ABB RobotStudio station: Pallet_Project.rspag

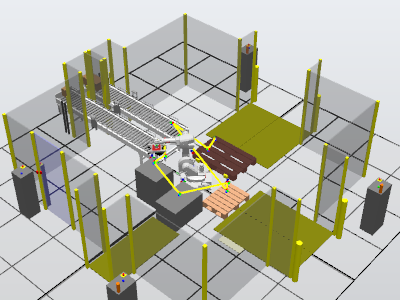
--- station ---
Station Pallet_Project (saved by RobotStudio 25.2.11220.0)
Controller Controler
  mechanical unit ROB_1: IRB1600_10_145__02, 6 joints, base frame (0, 0, 0) mm, rotated rx 0 ry 0 rz 135 deg
Layout (positions relative to the parent item):
  - IRB1600_10_145__02 [mechanism, from %ABB.RobotStudio.Models.IRB1600%\IRB1600_10_145_G_02.rslib] at (0, 0, 0) mm, rotated rx 0 ry 0 rz 135 deg; joint values [0, 0, 0, 0, 1.5708, 0] (rad or m)
  - Half EPAL [part] at (-400, -600, 0) mm, rotated rx 0 ry 0 rz -90 deg, size 600 x 800 x 144 mm
  - ConveyorBox1 [part, from %ABB.RobotStudio.Models.Conveyors%\Conveyor Guide 400.rslib] at (150, 3660, 0) mm, rotated rx 0 ry 0 rz -90 deg
  - ConveyorBox2 [part, from %ABB.RobotStudio.Models.Conveyors%\Conveyor Guide 400.rslib] at (-550, 3660, 0) mm, rotated rx 0 ry 0 rz -90 deg
  - PalletizingVacuumTool [mechanism] at (-530.33, 530.33, 1121.5) mm, rotated rx 180 ry 0 rz -45 deg
      TCP toolVacuum at (0, 0, 175) mm
      links: PalletizingVacuumTool
  - Box1 [part] at (338.5, 3410, 868) mm, size 249 x 499 x 200 mm
  - Box2 [part] at (-353.5, 3575, 868) mm, size 129 x 129 x 200 mm
  - EuroPallet [part, from Components\EuroPalletWood.rslib] at (1400, -600, 0) mm, rotated rx 0 ry 0 rz 90 deg
  - StackingTable [part], size 500 x 600 x 770 mm
  - LinerStand [part], size 800 x 540 x 500 mm
  - SC_Conveyor1 [smart component]
      signals: DO BoxArrived, DI EuroPalletReplaced, DO EuroPalletReplacedOut, DI EuroPalletFull
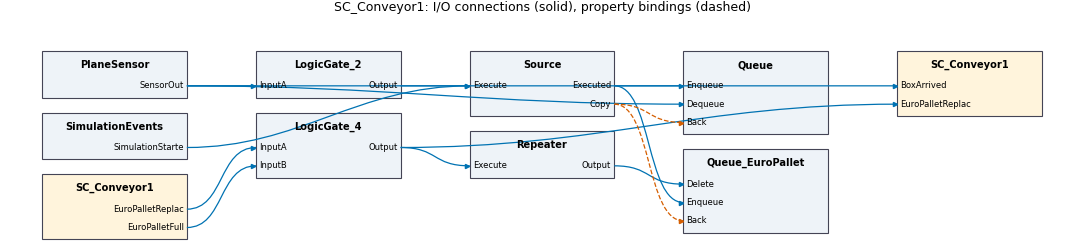
      connections:
        Source.Executed -> Queue.Enqueue
        PlaneSensor.SensorOut -> Queue.Dequeue
        PlaneSensor.SensorOut -> SC_Conveyor1.BoxArrived
        PlaneSensor.SensorOut -> LogicGate_2.InputA
        LogicGate_2.Output -> Source.Execute
        SimulationEvents.SimulationStarted -> Source.Execute
        SC_Conveyor1.EuroPalletReplaced -> LogicGate_4.InputA
        SC_Conveyor1.EuroPalletFull -> LogicGate_4.InputB
        LogicGate_4.Output -> SC_Conveyor1.EuroPalletReplacedOut
        LogicGate_4.Output -> Repeater.Execute
        Repeater.Output -> Queue_EuroPallet.Delete
        Source.Executed -> Queue_EuroPallet.Enqueue
        Source.Copy => Queue.Back
        Source.Copy => Queue_EuroPallet.Back
    - Source [smart component, from Components\Source.rslib]
        properties: Source=Box1; Copy=(none); Parent=(none); Position=[0.3385 3.39 0.868]; Orientation=[0 0 0]; Transient=true; PhysicsBehavior=-1
    - Queue [smart component, from Components\Queue.rslib]
        properties: Back=(none); Front=(none); Queue={70ca05b0-7144-4f49-83d8-d915b94a0a02};{7705e30e-55ab-4cc9-9220-690ff83121bf};{02bf6a2a-9363-4f0e-8f48-ba3ac55a3133};{2a754624-700a-40ce-a7f5-ac92a5654210};{9528570a-eb81-4ef3-89d0-eb89feb3dc99};{56097831-269e-4b26-b9dc-fc2a065cc4d2};{84102578-6d50-4318-bba9-f08da63948c5};{ab344251-b794-483f-853d-2cd57e9333d1};{43a68e49-bc40-4bf4-a0b0-52db603239fa};{90f7df2a-bd47-43a1-93ae-0975fdea56be};{8df4c4d2-3a0e-4db8-a3f9-2112c5fdeae1};{a6db4b97-f991-4390-b4fd-8137cccb983c};{ac275fb4-aa41-4d4d-8111-4fbb0763e808}; NumberOfObjects=1
    - LinearMover [smart component, from Components\LinearMover.rslib]
        properties: Object=Queue; Direction=[0 -0.001 0]; Speed=0.25; Reference=Global; ReferenceObject=(none)
    - PlaneSensor [smart component, from Components\PlaneSensor.rslib]
        properties: Origin=[0.1885 0.675 0.788]; Axis1=[0.3 0 0]; Axis2=[0 0 0.01]; Tag=(none); SenseMultiple=false; SensedPart=(none)
      - _sensorPart_ [part], size 300 x 0 x 10 mm
    - LogicGate_2 [smart component, from Components\LogicGate.rslib]
        properties: Operator=NOT; Delay=0
    - SimulationEvents [smart component, from Components\SimulationEvents.rslib]
    - Queue_EuroPallet [smart component, from Components\Queue.rslib]
        properties: Back=(none); Front=(none); Queue=; NumberOfObjects=0
    - LogicGate_4 [smart component, from Components\LogicGate.rslib]
        properties: Operator=AND; Delay=0
    - Repeater [smart component, from Components\Repeater.rslib]
        properties: Count=12
  - SC_Gripper [smart component]
      signals: DI Grip
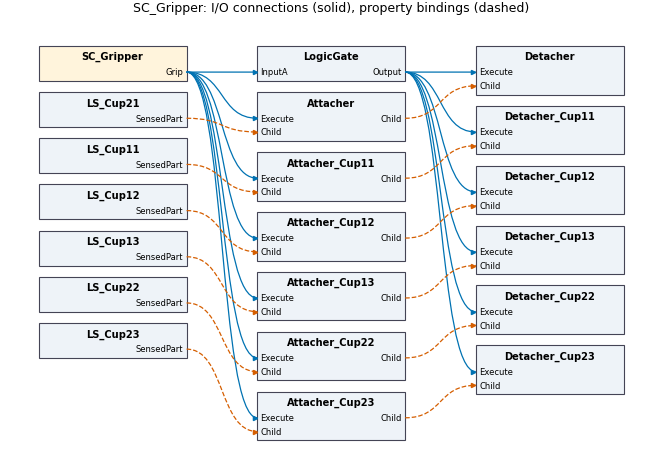
      connections:
        SC_Gripper.Grip -> Attacher.Execute
        SC_Gripper.Grip -> LogicGate.InputA
        LogicGate.Output -> Detacher.Execute
        SC_Gripper.Grip -> Attacher_Cup11.Execute
        LogicGate.Output -> Detacher_Cup11.Execute
        SC_Gripper.Grip -> Attacher_Cup12.Execute
        LogicGate.Output -> Detacher_Cup12.Execute
        SC_Gripper.Grip -> Attacher_Cup13.Execute
        LogicGate.Output -> Detacher_Cup13.Execute
        SC_Gripper.Grip -> Attacher_Cup22.Execute
        LogicGate.Output -> Detacher_Cup22.Execute
        SC_Gripper.Grip -> Attacher_Cup23.Execute
        LogicGate.Output -> Detacher_Cup23.Execute
        LS_Cup21.SensedPart => Attacher.Child
        Attacher.Child => Detacher.Child
        LS_Cup11.SensedPart => Attacher_Cup11.Child
        Attacher_Cup11.Child => Detacher_Cup11.Child
        LS_Cup12.SensedPart => Attacher_Cup12.Child
        Attacher_Cup12.Child => Detacher_Cup12.Child
        LS_Cup13.SensedPart => Attacher_Cup13.Child
        Attacher_Cup13.Child => Detacher_Cup13.Child
        LS_Cup22.SensedPart => Attacher_Cup22.Child
        Attacher_Cup22.Child => Detacher_Cup22.Child
        LS_Cup23.SensedPart => Attacher_Cup23.Child
        Attacher_Cup23.Child => Detacher_Cup23.Child
    - LS_Cup21 [smart component, from Components\LineSensor.rslib] at (0, 0, 0) mm
        properties: Start=[-0.597509982704304 0.689429996191639 0.956499992313755]; End=[-0.597509981617333 0.689429995104668 0.924499992313755]; Length=0.032; Radius=0.00331491712707182; Tag=(none); SenseMultiple=false; SensedPart=(none); SensedPoint=[0 0 0]
      - _sensorPart_ [part], size 6.4 x 6.4 x 32 mm
    - Attacher [smart component, from Components\Attacher.rslib]
        properties: Parent=PalletizingVacuumTool; Flange=0; Child=(none); Mount=false; Offset=[0 0 0]; Orientation=[0 0 0]
    - Detacher [smart component, from Components\Detacher.rslib]
        properties: Child=(none); KeepPosition=true
    - LogicGate [smart component, from Components\LogicGate.rslib]
        properties: Operator=NOT; Delay=0
    - LS_Cup11 [smart component, from Components\LineSensor.rslib]
        properties: Start=[-0.68943 0.59751 0.9565]; End=[-0.68943 0.59751 0.9245]; Length=0.032; Radius=0.00331; Tag=(none); SenseMultiple=false; SensedPart=(none); SensedPoint=[0 0 0]
      - _sensorPart_ [part], size 6.6 x 6.6 x 32 mm
    - LS_Cup12 [smart component, from Components\LineSensor.rslib]
        properties: Start=[-0.57629 0.48437 0.9565]; End=[-0.57629 0.48437 0.9245]; Length=0.032; Radius=0.00331; Tag=(none); SenseMultiple=false; SensedPart=(none); SensedPoint=[0 0 0]
      - _sensorPart_ [part], size 6.6 x 6.6 x 32 mm
    - LS_Cup13 [smart component, from Components\LineSensor.rslib]
        properties: Start=[-0.46315 0.37123 0.9565]; End=[-0.46315 0.37123 0.9245]; Length=0.032; Radius=0.00331; Tag=(none); SenseMultiple=false; SensedPart=(none); SensedPoint=[0 0 0]
      - _sensorPart_ [part], size 6.6 x 6.6 x 32 mm
    - LS_Cup22 [smart component, from Components\LineSensor.rslib]
        properties: Start=[-0.48437 0.57629 0.9565]; End=[-0.48437 0.57629 0.9245]; Length=0.032; Radius=0.00331; Tag=(none); SenseMultiple=false; SensedPart=(none); SensedPoint=[0 0 0]
      - _sensorPart_ [part], size 6.6 x 6.6 x 32 mm
    - LS_Cup23 [smart component, from Components\LineSensor.rslib]
        properties: Start=[-0.37123 0.46315 0.9565]; End=[-0.37123 0.46315 0.9245]; Length=0.032; Radius=0.00331; Tag=(none); SenseMultiple=false; SensedPart=(none); SensedPoint=[0 0 0]
      - _sensorPart_ [part], size 6.6 x 6.6 x 32 mm
    - Attacher_Cup11 [smart component, from Components\Attacher.rslib]
        properties: Parent=PalletizingVacuumTool; Flange=0; Child=(none); Mount=false; Offset=[0 0 0]; Orientation=[0 0 0]
    - Detacher_Cup11 [smart component, from Components\Detacher.rslib]
        properties: Child=(none); KeepPosition=true
    - Attacher_Cup12 [smart component, from Components\Attacher.rslib]
        properties: Parent=PalletizingVacuumTool; Flange=0; Child=(none); Mount=false; Offset=[0 0 0]; Orientation=[0 0 0]
    - Detacher_Cup12 [smart component, from Components\Detacher.rslib]
        properties: Child=(none); KeepPosition=true
    - Attacher_Cup13 [smart component, from Components\Attacher.rslib]
        properties: Parent=PalletizingVacuumTool; Flange=0; Child=(none); Mount=false; Offset=[0 0 0]; Orientation=[0 0 0]
    - Detacher_Cup13 [smart component, from Components\Detacher.rslib]
        properties: Child=(none); KeepPosition=true
    - Attacher_Cup22 [smart component, from Components\Attacher.rslib]
        properties: Parent=PalletizingVacuumTool; Flange=0; Child=(none); Mount=false; Offset=[0 0 0]; Orientation=[0 0 0]
    - Detacher_Cup22 [smart component, from Components\Detacher.rslib]
        properties: Child=(none); KeepPosition=true
    - Attacher_Cup23 [smart component, from Components\Attacher.rslib]
        properties: Parent=PalletizingVacuumTool; Flange=0; Child=(none); Mount=false; Offset=[0 0 0]; Orientation=[0 0 0]
    - Detacher_Cup23 [smart component, from Components\Detacher.rslib]
        properties: Child=(none); KeepPosition=true
  - SC_Conveyor2 [smart component]
      signals: DO BoxArrived, DI HalfPalletReplaced, DI HalfPalletFull, DO HalfPalletReplacedOut
      connections:
        Source.Executed -> Queue.Enqueue
        PlaneSensor.SensorOut -> Queue.Dequeue
        PlaneSensor.SensorOut -> SC_Conveyor2.BoxArrived
        PlaneSensor.SensorOut -> LogicGate.InputA
        SimulationEvents.SimulationStarted -> Source.Execute
        Source.Executed -> Queue_HalfPallet.Enqueue
        LogicGate.Output -> Source.Execute
        Repeater.Output -> Queue_HalfPallet.Delete
        SC_Conveyor2.HalfPalletReplaced -> LogicGate_5.InputA
        SC_Conveyor2.HalfPalletFull -> LogicGate_5.InputB
        LogicGate_5.Output -> Repeater.Execute
        LogicGate_5.Output -> SC_Conveyor2.HalfPalletReplacedOut
        Source.Copy => Queue.Back
        Source.Copy => Queue_HalfPallet.Back
    - Source [smart component, from Components\Source.rslib]
        properties: Source=Box2; Copy=(none); Parent=(none); Position=[-0.3535 3.575 0.868]; Orientation=[0 0 0]; Transient=true; PhysicsBehavior=-1
    - Queue [smart component, from Components\Queue.rslib]
        properties: Back=(none); Front=(none); Queue={648eb2a2-8d13-4a50-a9a9-4bb0657455f7};{41be35e7-4a03-4cb4-92d6-970da98b32eb};{4f5e8617-4ef4-4248-bc63-4e8ec75bf0fd};{9850fa1d-30e0-46cb-a9aa-89d687d5a572};{8673d542-8e4c-49b3-88b3-ba839af60b27};{121a61d2-9307-4f78-a061-101ab78a5607};{316e579a-2297-4da1-921e-c195e3c1eac9};{afd6ccd5-80c3-46f0-a33f-b3bd5f1b0761};{a691a1e4-6464-4329-bb8e-435514d80af1};{358ac2eb-a4d6-456f-aa39-476db23d4f48}; NumberOfObjects=1
    - LinearMover [smart component, from Components\LinearMover.rslib]
        properties: Object=Queue; Direction=[0 -0.001 0]; Speed=0.25; Reference=Global; ReferenceObject=(none)
    - PlaneSensor [smart component, from Components\PlaneSensor.rslib]
        properties: Origin=[-0.5035 0.675 0.788]; Axis1=[0.3 0 0]; Axis2=[0 0 0.01]; Tag=(none); SenseMultiple=false; SensedPart=(none)
      - _sensorPart_ [part], size 300 x 0 x 10 mm
    - LogicGate [smart component, from Components\LogicGate.rslib]
        properties: Operator=NOT; Delay=0
    - SimulationEvents [smart component, from Components\SimulationEvents.rslib]
    - Queue_HalfPallet [smart component, from Components\Queue.rslib]
        properties: Back=(none); Front=(none); Queue={f5edb1ce-3bf5-426a-a389-0b0047efa949};{5ce0816a-b692-43c6-82f7-492eb3fc1c7c};{ad3ef4b5-2c59-4daa-9658-0c77e5efb67d};{c9c476d0-74ff-4b18-bfb3-2d6c852b8493};{1bf865c6-1649-4319-b5ff-cd81faaa6069};{f626778c-15a6-4059-b27a-7c8f9da4f34f};{a60dd0dd-490e-48fe-bb32-16f415136b44};{4ec9b3b2-e4a8-4d14-aea0-9552a35d2afd};{38bc6a68-8d9e-44a7-a5f0-badb214ea710};{f9543542-377a-43f1-9613-018dced76680};{486b4c2f-b225-4486-b430-5ab7d813c599};{7da52d9e-9053-4b1a-839c-0aedc5495cc7};{c2400356-fde5-4523-9dc7-d26788098951};{75099568-1fe6-4c34-8328-63fd42144c3b};{8ca6c374-2d39-4938-8324-38c48ae4f51d};{f3c160ab-6f5f-460b-8b54-c2c3b0bc175f};{1c289510-9a29-4e1c-b603-54b7a0027260};{d39da69b-e59a-4ace-85a5-bba54583b01c};{bc328c62-4bf3-4a57-965c-0c93e0ee296d};{60f4dcb3-d366-4d0b-b05a-5b2073fcd9e8};{44334a49-cf52-4d95-9964-3bb568ce732d};{f9240695-1965-47e5-bcd4-644ec5904899};{72a970fd-f238-4ac5-b811-00686975bc20};{bd297b2a-4ad7-44fa-87c8-1ac40b0d2fbf};{3dafa88d-62b0-429f-9c75-c8c7bde09fc6};{a7d8f176-4e9d-4819-8805-982bee0c310d};{72ae6bb6-3373-4f60-a321-dfdc0981c562};{fff16105-3d56-4b21-a888-399904fd95d4};{56e4abf9-acd4-4a00-b067-52a58200d221};{2eb8ae55-b553-4f83-b65d-07c27c701dd6};{dfb05241-1220-45e8-b584-1559777c0125};{49a2c23a-27ea-4b0b-af5c-f9d01014f642};{0adfb5d7-4fd0-41be-8361-c42c9d28ca51};{8cf74624-f46b-49ca-a524-038ddb88ba0f};{bde2cdc4-b3e4-48fe-8333-d64185b5a8e7};{d17564c2-89d4-4b4f-8596-5dca9165a286};{6fec26e7-cb1b-4d74-b4a6-8ed7a2eb81a6};{e04d8697-cc19-4df5-b7fa-dff41516820c};{134714af-70a5-49a3-8b99-ea847d1ef329};{23aa8eff-aaeb-4079-b6e6-9fe5f0b7799c};{0091a76d-e23e-4382-9bf3-a427b049953f};{fdc2abc9-40b2-462e-8472-b1d156765a68};{8dc86a38-8dcf-454b-a79a-3f5e6d46a581};{f9226736-fe9f-4ce5-82b5-97fc8f487c87};{8d0584df-2d5d-4d5a-bd5b-c865cb85c145};{fef2818e-b6b9-47fe-bf8a-83543bb000b1}; NumberOfObjects=7
    - Repeater [smart component, from Components\Repeater.rslib]
        properties: Count=72
    - LogicGate_5 [smart component, from Components\LogicGate.rslib]
        properties: Operator=AND; Delay=0
  - Liner_01 [part] at (-900, -2000, 0) mm, size 800 x 540 x 10 mm
  - SC_Liners [smart component]
      signals: DI LinersRefilled, DI LinerStackEmpty, DI PalletReplaced, DO LinersRefilledOut
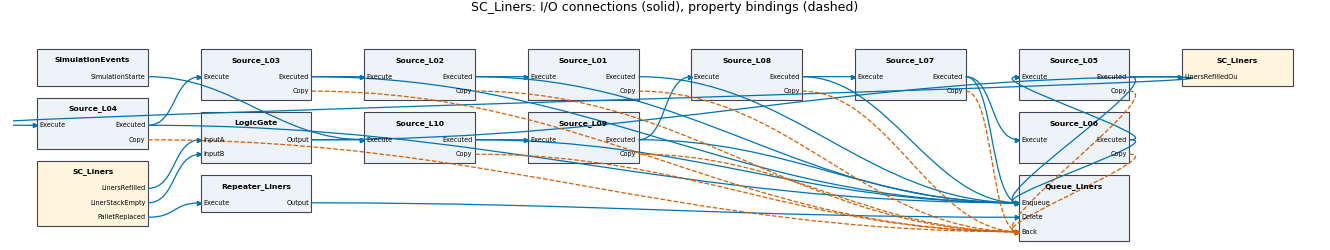
      connections:
        SimulationEvents.SimulationStarted -> Source_L10.Execute
        Source_L10.Executed -> Queue_Liners.Enqueue
        Source_L10.Executed -> Source_L09.Execute
        Source_L09.Executed -> Queue_Liners.Enqueue
        Source_L09.Executed -> Source_L08.Execute
        Source_L08.Executed -> Queue_Liners.Enqueue
        Source_L08.Executed -> Source_L07.Execute
        Source_L07.Executed -> Queue_Liners.Enqueue
        Source_L07.Executed -> Source_L06.Execute
        Source_L06.Executed -> Queue_Liners.Enqueue
        Source_L06.Executed -> Source_L05.Execute
        Source_L05.Executed -> Queue_Liners.Enqueue
        Source_L05.Executed -> Source_L04.Execute
        Source_L04.Executed -> Queue_Liners.Enqueue
        Source_L04.Executed -> Source_L03.Execute
        Source_L03.Executed -> Queue_Liners.Enqueue
        Source_L03.Executed -> Source_L02.Execute
        Source_L02.Executed -> Queue_Liners.Enqueue
        Source_L02.Executed -> Source_L01.Execute
        Source_L01.Executed -> Queue_Liners.Enqueue
        SC_Liners.LinersRefilled -> LogicGate.InputA
        SC_Liners.LinerStackEmpty -> LogicGate.InputB
        LogicGate.Output -> SC_Liners.LinersRefilledOut
        LogicGate.Output -> Source_L10.Execute
        SC_Liners.PalletReplaced -> Repeater_Liners.Execute
        Repeater_Liners.Output -> Queue_Liners.Delete
        Source_L10.Copy => Queue_Liners.Back
        Source_L09.Copy => Queue_Liners.Back
        Source_L08.Copy => Queue_Liners.Back
        Source_L07.Copy => Queue_Liners.Back
        Source_L06.Copy => Queue_Liners.Back
        Source_L05.Copy => Queue_Liners.Back
        Source_L04.Copy => Queue_Liners.Back
        Source_L03.Copy => Queue_Liners.Back
        Source_L02.Copy => Queue_Liners.Back
        Source_L01.Copy => Queue_Liners.Back
    - Source_L10 [smart component, from Components\Source.rslib]
        properties: Source=Liner_01; Copy=(none); Parent=(none); Position=[-1.3 -0.7 0.59]; Orientation=[0 0 0]; Transient=true; PhysicsBehavior=-1
    - Source_L09 [smart component, from Components\Source.rslib]
        properties: Source=Liner_01; Copy=(none); Parent=(none); Position=[-1.3 -0.7 0.58]; Orientation=[0 0 0]; Transient=true; PhysicsBehavior=-1
    - Queue_Liners [smart component, from Components\Queue.rslib]
        properties: Back=(none); Front=(none); Queue={4b76874b-49d8-40e7-b1bf-01d8cc753daf};{f1bc3993-1843-4745-a916-cd233907ef8f}; NumberOfObjects=2
    - SimulationEvents [smart component, from Components\SimulationEvents.rslib]
    - Source_L08 [smart component, from Components\Source.rslib]
        properties: Source=Liner_01; Copy=(none); Parent=(none); Position=[-1.3 -0.7 0.57]; Orientation=[0 0 0]; Transient=true; PhysicsBehavior=-1
    - Source_L07 [smart component, from Components\Source.rslib]
        properties: Source=Liner_01; Copy=(none); Parent=(none); Position=[-1.3 -0.7 0.56]; Orientation=[0 0 0]; Transient=true; PhysicsBehavior=-1
    - Source_L06 [smart component, from Components\Source.rslib]
        properties: Source=Liner_01; Copy=(none); Parent=(none); Position=[-1.3 -0.7 0.55]; Orientation=[0 0 0]; Transient=true; PhysicsBehavior=-1
    - Source_L05 [smart component, from Components\Source.rslib]
        properties: Source=Liner_01; Copy=(none); Parent=(none); Position=[-1.3 -0.7 0.54]; Orientation=[0 0 0]; Transient=true; PhysicsBehavior=-1
    - Source_L04 [smart component, from Components\Source.rslib]
        properties: Source=Liner_01; Copy=(none); Parent=(none); Position=[-1.3 -0.7 0.53]; Orientation=[0 0 0]; Transient=true; PhysicsBehavior=-1
    - Source_L03 [smart component, from Components\Source.rslib]
        properties: Source=Liner_01; Copy=(none); Parent=(none); Position=[-1.3 -0.7 0.52]; Orientation=[0 0 0]; Transient=true; PhysicsBehavior=-1
    - Source_L02 [smart component, from Components\Source.rslib]
        properties: Source=Liner_01; Copy=(none); Parent=(none); Position=[-1.3 -0.7 0.51]; Orientation=[0 0 0]; Transient=true; PhysicsBehavior=-1
    - Source_L01 [smart component, from Components\Source.rslib]
        properties: Source=Liner_01; Copy=(none); Parent=(none); Position=[-1.3 -0.7 0.5]; Orientation=[0 0 0]; Transient=true; PhysicsBehavior=-1
    - LogicGate [smart component, from Components\LogicGate.rslib]
        properties: Operator=AND; Delay=0
    - Repeater_Liners [smart component, from Components\Repeater.rslib]
        properties: Count=2
  - Door_Maintenance [part], size 20 x 800 x 2000 mm
  - LightCurtain_EuroPallet_Emitter [part], size 50 x 50 x 2000 mm
  - LightCurtain_EuroPallet_Receiver [part], size 50 x 50 x 2000 mm
  - LightCurtain_HalfPallet_Emitter [part], size 50 x 50 x 2000 mm
  - LightCurtain_HalfPallet_Receiver [part], size 50 x 50 x 2000 mm
  - LightCurtain_LinerBay_Emitter [part], size 50 x 50 x 2000 mm
  - LightCurtain_LinerBay_Receiver [part], size 50 x 50 x 2000 mm
  - LightCurtain_Conv1_Emitter [part], size 50 x 50 x 450 mm
  - LightCurtain_Conv1_Receiver [part], size 50 x 50 x 450 mm
  - LightCurtain_Conv2_Emitter [part], size 50 x 50 x 450 mm
  - LightCurtain_Conv2_Receiver [part], size 50 x 50 x 450 mm
  - MutingSensor_Conv1_A [part], size 30 x 30 x 900 mm
  - MutingSensor_Conv1_B [part], size 30 x 30 x 900 mm
  - MutingSensor_Conv2_A [part], size 30 x 30 x 900 mm
  - MutingSensor_Conv2_B [part], size 30 x 30 x 900 mm
  - SafetyMat_EuroPallet [part], size 1650 x 1800 x 15 mm
  - SafetyMat_HalfPallet [part], size 1500 x 1850 x 15 mm
  - SafetyMat_LinerBay [part], size 1750 x 740 x 15 mm
  - PalletStop_Euro_1 [part], size 40 x 100 x 80 mm
  - PalletStop_Euro_2 [part], size 40 x 100 x 80 mm
  - PalletStop_Half_1 [part], size 100 x 40 x 80 mm
  - PalletStop_Half_2 [part], size 100 x 40 x 80 mm
  - OperatorStation_EuroPallet [part], size 400 x 300 x 1100 mm
  - OperatorStation_HalfPallet [part], size 400 x 300 x 1100 mm
  - OperatorStation_LinerBay [part], size 400 x 300 x 1100 mm
  - OperatorStation_General [part], size 400 x 300 x 1100 mm
  - OperatorStation_Door [part], size 300 x 300 x 1100 mm
  - EStopPost_Inside [part], size 100 x 100 x 1100 mm
  - IRC5_Cabinet [part], size 725 x 710 x 970 mm
  - DoorSensor_Eden_Actuator [part], size 30 x 40 x 60 mm
  - DoorSensor_Eden_Sensor [part], size 30 x 40 x 60 mm
  - EStopBase_EuroPallet [part], size 80 x 80 x 5 mm
  - EStopBase_HalfPallet [part], size 80 x 80 x 5 mm
  - EStopBase_LinerBay [part], size 80 x 80 x 5 mm
  - EStopBase_General [part], size 80 x 80 x 5 mm
  - EStopBase_Door [part], size 80 x 80 x 5 mm
  - EStopBase_Inside [part], size 80 x 80 x 5 mm
  - Bumper_EuroPallet_1 [part], size 114 x 114 x 1000 mm
  - Bumper_EuroPallet_2 [part], size 114 x 114 x 1000 mm
  - Bumper_HalfPallet_1 [part], size 114 x 114 x 1000 mm
  - Bumper_HalfPallet_2 [part], size 114 x 114 x 1000 mm
  - MutingLamp_Conv1 [part], size 60 x 60 x 100 mm
  - MutingLamp_Conv2 [part], size 60 x 60 x 100 mm
  - Lamp_EuroPalletFull [part], size 60 x 59.8 x 200 mm
  - Lamp_HalfPalletFull [part], size 60 x 59.8 x 200 mm
  - Lamp_LinerStackEmpty [part], size 60 x 59.8 x 200 mm
  - Button_EuroPalletReplaced [part], size 40 x 39.9 x 20 mm
  - Button_HalfPalletReplaced [part], size 40 x 39.9 x 20 mm
  - Button_LinersRefilled [part], size 40 x 39.9 x 20 mm
  - ResetButton_EuroPallet [part], size 40 x 39.9 x 20 mm
  - ResetButton_HalfPallet [part], size 40 x 39.9 x 20 mm
  - ResetButton_LinerBay [part], size 40 x 39.9 x 20 mm
  - ResetButton_Door [part], size 40 x 39.9 x 20 mm
  - EStop_EuroPallet [part], size 40 x 40 x 30 mm
  - EStop_HalfPallet [part], size 40 x 40 x 30 mm
  - EStop_LinerBay [part], size 40 x 40 x 30 mm
  - EStop_General [part], size 40 x 40 x 30 mm
  - EStop_Door [part], size 40 x 40 x 30 mm
  - EStop_Inside [part], size 40 x 40 x 30 mm
  - Safety_Fence [graphiccomponentgroup]
    - Fence_Corridor_Euro_1 [part], size 500 x 20 x 2000 mm
    - Fence_Corridor_Euro_2 [part], size 500 x 20 x 2000 mm
    - Fence_Corridor_Half_1 [part], size 20 x 500 x 2000 mm
    - Fence_Corridor_Half_2 [part], size 20 x 500 x 2000 mm
    - Fence_Corridor_Liner_1 [part], size 500 x 20 x 2000 mm
    - Fence_Corridor_Liner_2 [part], size 500 x 20 x 2000 mm
    - Fence_Panel_E1 [part], size 20 x 1650 x 2000 mm
    - Fence_Panel_E2 [part], size 20 x 1650 x 2000 mm
    - Fence_Panel_N1 [part], size 1931.5 x 20 x 2000 mm
    - Fence_Panel_N2 [part], size 162 x 20 x 2000 mm
    - Fence_Panel_N3 [part], size 1946.5 x 20 x 2000 mm
    - Fence_Panel_S1 [part], size 1800 x 20 x 2000 mm
    - Fence_Panel_S2 [part], size 1800 x 20 x 2000 mm
    - Fence_Panel_W1 [part], size 20 x 1750 x 2000 mm
    - Fence_Panel_W2 [part], size 20 x 960 x 2000 mm
    - Fence_Panel_W3 [part], size 20 x 850 x 2000 mm
    - Fence_Post_01 [part], size 60 x 60 x 2000 mm
    - Fence_Post_02 [part], size 60 x 60 x 2000 mm
    - Fence_Post_03 [part], size 60 x 60 x 2000 mm
    - Fence_Post_04 [part], size 60 x 60 x 2000 mm
    - Fence_Post_05 [part], size 60 x 60 x 2000 mm
    - Fence_Post_06 [part], size 60 x 60 x 2000 mm
    - Fence_Post_07 [part], size 60 x 60 x 2000 mm
    - Fence_Post_08 [part], size 60 x 60 x 2000 mm
    - Fence_Post_09 [part], size 60 x 60 x 2000 mm
    - Fence_Post_10 [part], size 60 x 60 x 2000 mm
    - Fence_Post_11 [part], size 60 x 60 x 2000 mm
    - Fence_Post_12 [part], size 60 x 60 x 2000 mm
    - Fence_Post_13 [part], size 60 x 60 x 2000 mm
    - Fence_Post_14 [part], size 60 x 60 x 2000 mm
    - Fence_Post_15 [part], size 60 x 60 x 2000 mm
    - Fence_Post_16 [part], size 60 x 60 x 2000 mm
    - Fence_Post_17 [part], size 60 x 60 x 2000 mm
    - Fence_Post_18 [part], size 60 x 60 x 2000 mm
    - Fence_Post_19 [part], size 60 x 60 x 2000 mm
    - Fence_Post_20 [part], size 60 x 60 x 2000 mm
    - Fence_Tunnel_Conv1_1 [part], size 20 x 500 x 2000 mm
    - Fence_Tunnel_Conv1_2 [part], size 20 x 500 x 2000 mm
    - Fence_Tunnel_Conv1_Low [part], size 530 x 20 x 700 mm
    - Fence_Tunnel_Conv1_Top [part], size 530 x 20 x 980 mm
    - Fence_Tunnel_Conv2_1 [part], size 20 x 500 x 2000 mm
    - Fence_Tunnel_Conv2_2 [part], size 20 x 500 x 2000 mm
    - Fence_Tunnel_Conv2_Low [part], size 530 x 20 x 700 mm
    - Fence_Tunnel_Conv2_Top [part], size 530 x 20 x 980 mm
Attachment: PalletizingVacuumTool is attached to IRB1600_10_145__02 / Link6
Attachment: LS_Cup21 is attached to PalletizingVacuumTool / PalletizingVacuumTool
Attachment: LS_Cup12 is attached to PalletizingVacuumTool / PalletizingVacuumTool
Attachment: LS_Cup13 is attached to PalletizingVacuumTool / PalletizingVacuumTool
Attachment: LS_Cup22 is attached to PalletizingVacuumTool / PalletizingVacuumTool
Attachment: LS_Cup23 is attached to PalletizingVacuumTool / PalletizingVacuumTool
Attachment: LS_Cup11 is attached to PalletizingVacuumTool / PalletizingVacuumTool
Collision set Conjunto de colisión_1: IRB1600_10_145__02, PalletizingVacuumTool against ConveyorBox1, ConveyorBox2, EuroPallet, Half EPAL, LinerStand, StackingTable, near miss 0.05 m
Station logic (signal -> signal, property => property):
  SC_Conveyor1.BoxArrived -> Controler.DI_Box1Arrived
  Controler.DO_Cup21 -> SC_Gripper.Grip
  SC_Conveyor2.BoxArrived -> Controler.DI_Box2Arrived
  SC_Conveyor1.EuroPalletReplacedOut -> Controler.DI_EuroPalletReplaced
  Controler.DO_EuroPalletFull -> SC_Conveyor1.EuroPalletFull
  Controler.DO_HalfPalletFull -> SC_Conveyor2.HalfPalletFull
  SC_Conveyor2.HalfPalletReplacedOut -> Controler.DI_HalfPalletReplaced
  Controler.DO_LinerStackEmpty -> SC_Liners.LinerStackEmpty
  SC_Liners.LinersRefilledOut -> Controler.DI_LinersRefilled
  SC_Conveyor2.HalfPalletReplacedOut -> SC_Liners.PalletReplaced
Targets, tools, work objects and paths stored in the station and not in the controller backup, written as RAPID:
! task T_ROB1
MODULE PalletProgram
  PROC Path_10()
    MoveL PickConveyor2,v1000,z100,toolVacuum\WObj:=wobjConveyor2;
    MoveL PlaceTable,v1000,z100,toolVacuum\WObj:=wobjTable;
    MoveL PickTableStack,v1000,z100,toolVacuum\WObj:=wobjTable;
    MoveL PickLiner,v1000,z100,toolVacuum\WObj:=wobjLinerStack;
    MoveL PlaceHalfPallet,v1000,z100,toolVacuum\WObj:=wobjHalfPallet;
    MoveL PlaceLiner,v1000,z100,toolVacuum\WObj:=wobjHalfPallet;
    MoveL PickConveyor1,v1000,z100,toolVacuum\WObj:=wobjConveyor1;
    MoveL PlaceEuroRow2,v1000,z100,toolVacuum\WObj:=wobjEuroPallet;
    MoveL PlaceEuroRow4,v1000,z100,toolVacuum\WObj:=wobjEuroPallet;
  ENDPROC
ENDMODULE


--- Controller Data/Controler/RAPID/TASK1/PROGMOD/CalibData.mod ---
MODULE CalibData
    ! Calibration data: work objects, tool and loads (mm, kg).
    ! Work objects are given in the world frame (wobj0 = world, not the robot base).

    !-----------------------------------------------------------------------
    ! Work objects and tool
    !-----------------------------------------------------------------------
    ! Euro pallet (1200x800): origin at the corner nearest the robot and conveyor 1, on top of the
    ! pallet (z 144). X along the long side, away from the conveyors; Y away from the robot
    TASK PERS wobjdata wobjEuroPallet:=[FALSE,TRUE,"",[[600,600,144],[0.707106781,0,0,-0.707106781]],[[0,0,0],[1,0,0,0]]];
    ! Half pallet (800x600): origin at the corner nearest the robot and the Euro pallet, on top of the
    ! pallet (z 144). X along the long side, towards the liner stand; Y away from the robot
    TASK PERS wobjdata wobjHalfPallet:=[FALSE,TRUE,"",[[400,-600,144],[0,0,0,1]],[[0,0,0],[1,0,0,0]]];
    ! Conveyor 1 (Euro pallet side): origin at the end next to the robot, centred on the belt (z 768).
    ! X along the conveyor, against the flow; Y towards conveyor 2
    TASK PERS wobjdata wobjConveyor1:=[FALSE,TRUE,"",[[338.5,670,768],[0.707106781,0,0,0.707106781]],[[0,0,0],[1,0,0,0]]];
    ! Conveyor 2 (table side): same as conveyor 1. X against the flow; Y away from conveyor 1
    TASK PERS wobjdata wobjConveyor2:=[FALSE,TRUE,"",[[-353.5,670,768],[0.707106781,0,0,0.707106781]],[[0,0,0],[1,0,0,0]]];
    ! Stacking table: origin at the corner next to the end of conveyor 2, on the table top (z 770).
    ! X away from conveyor 2; Y in the direction the boxes travel on the conveyors.
    ! oframe (55,170) centres the 3x2 block on the table
    TASK PERS wobjdata wobjTable:=[FALSE,TRUE,"",[[-600,600,770],[0,0,0,1]],[[55,170,0],[1,0,0,0]]];
    ! Liner stand: origin at the corner nearest the robot and the half pallet, on top of the stand
    ! (z 500, base of the liner stack). X along the long side (800 mm liner), away from the half pallet;
    ! Y away from the robot
    TASK PERS wobjdata wobjLinerStack:=[FALSE,TRUE,"",[[-500,-160,500],[0,0,0,1]],[[0,0,0],[1,0,0,0]]];
    ! toolVacuum: TCP on the cup faces, 175 mm from the flange, at the centre of the 6 cups
    ! Mass estimated from the measured parts in aluminium (2700 kg/m3), with the column as a tube
    ! and the grey plate hollow (5 mm walls): 4.65 kg, rounded up to 4.7 kg. CoG on the tool axis,
    ! 100 mm from the flange (tool0). Solid as drawn it would be 9.6 kg: more than the 10 kg payload
    ! of the robot together with the 2.4 kg block. Inertia about the CoG, from the same parts
    ! (cylinders, plates and 6 cups as point masses of 0.05 kg)
    TASK PERS tooldata toolVacuum:=[TRUE,[[0,0,175],[1,0,0,0]],[4.7,[0,0,100],[1,0,0,0],0.0274,0.0462,0.0605]];

    !-----------------------------------------------------------------------
    ! Load data
    !-----------------------------------------------------------------------
    ! Payloads: CoG relative to the TCP of toolVacuum. Inertia about the CoG of the load, as a solid
    ! box: Ix = m(b2+c2)/12, Iy = m(a2+c2)/12, Iz = m(a2+b2)/12 (a, b, c = size along tool X, Y, Z)
    ! Box 1: 500 x 250 x 200 mm (long side along the tool X), 2 kg
    TASK PERS loaddata loadBox1:=[2,[0,0,100],[1,0,0,0],0.0171,0.0483,0.0521];
    ! Box 2: 130 x 130 x 200 mm, 0.4 kg. Picked with one corner cup (Cup21, x=-160, y=-100 from
    ! the TCP): the CoG is under that cup
    TASK PERS loaddata loadBox2:=[0.4,[-160,-100,100],[1,0,0,0],0.0019,0.0019,0.0011];
    ! 3x2 block of box 2: 390 x 260 x 200 mm (3 boxes along the tool X), 6 x 0.4 kg
    TASK PERS loaddata loadBox2Stack:=[2.4,[0,0,100],[1,0,0,0],0.0215,0.0384,0.0439];
    ! Liner: corrugated cardboard, 0.8 x 0.54 x 0.01 m3 x 120 kg/m3 = 0.52 kg (800 mm along the tool X)
    TASK PERS loaddata loadLiner:=[0.52,[0,0,5],[1,0,0,0],0.0126,0.0277,0.0404];
ENDMODULE

--- Controller Data/Controler/RAPID/TASK1/PROGMOD/PalletProgram.mod ---
MODULE PalletProgram

    !***********************************************************************
    ! Industrial Robotics and Offline Programming G1F - University of Skovde
    ! Offline programming project: Pallet Project - Group 2 (JMPM)
    ! Authors: Peru Mendivil and Joaquin Moreno
    ! Robot :   ABB IRB 1600-10/1.45, IRC5 RobotWare 6.13.02 (RobotStudio 2025)
    ! Tool  :   toolVacuum, vacuum gripper with 6 cups (one valve per cup)
    ! Date:    2026-10-30
    !
    ! The robot palletizes two products coming on two conveyors.
    ! Box 1 goes from conveyor 1 to the Euro pallet: 4-2 pattern,
    ! 2 layers (12 boxes). Box 2 goes from conveyor 2 to the stacking
    ! table, where a 3x2 block is formed. The block is then moved to the
    ! half pallet: 2x2 blocks per layer, 3 layers (72 boxes), with a liner
    ! after layers 1 and 2. When both conveyors have a box, the robot
    ! alternates box 1 and box 2. A full pallet is replaced by the operator
    ! from outside the fence, and the robot keeps working with the other
    ! product. With the half pallet full, one block can still be finished
    ! on the table, and it waits there. If the liner stack is empty, the
    ! robot keeps working until a liner is needed; then box 2 waits until
    ! the operator refills the stack.
    !
    ! Structure: Main is a state machine (grafcet). It initialises the
    ! signals and then decides each cycle which box to handle, from the
    ! conveyor sensors, the full-pallet flags and the last box handled.
    ! Each product has its own routine with a finite-state machine for
    ! the place positions. Every place position is calculated with Offs
    ! from one base target per station. ApproachPoint does every
    ! pick/place: approach, vacuum on/off and GripLoad. Work objects,
    ! tool and loads are in the module CalibData.
    ! The operator buttons (pallet replaced, liners refilled) are read
    ! with interrupts (TRAP), so a short press is never lost.
    !
    ! Naming: VAR, PERS and parameters in camelCase (can change);
    ! CONST, PROC, FUNC and MODULE in PascalCase (fixed).
    !***********************************************************************

    !-----------------------------------------------------------------------
    ! Base targets
    !-----------------------------------------------------------------------
    CONST jointtarget Home:=[[0,0,0,0,90,0],[9E+09,9E+09,9E+09,9E+09,9E+09,9E+09]];

    ! Box 1
    CONST robtarget PickConveyor1:=[[249.5,0,200],[0,0,1,0],[0,0,0,0],[9E+09,9E+09,9E+09,9E+09,9E+09,9E+09]];
    CONST robtarget PlaceEuroRow4:=[[225,525,200],[0,-0.707106781,0.707106781,0],[-2,0,0,0],[9E+09,9E+09,9E+09,9E+09,9E+09,9E+09]];
    CONST robtarget PlaceEuroRow2:=[[350,150,200],[0,1,0,0],[-2,0,-1,0],[9E+09,9E+09,9E+09,9E+09,9E+09,9E+09]];

    ! Box 2
    CONST robtarget PickConveyor2:=[[-35.5,-160,200],[0,-0.707106781,0.707106781,0],[0,0,0,0],[9E+09,9E+09,9E+09,9E+09,9E+09,9E+09]];
    CONST robtarget PlaceTable:=[[-95,165,200],[0,0,1,0],[0,0,0,0],[9E+09,9E+09,9E+09,9E+09,9E+09,9E+09]];
    CONST robtarget PickTableStack:=[[195,130,200],[0,0,1,0],[0,0,0,0],[9E+09,9E+09,9E+09,9E+09,9E+09,9E+09]];
    CONST robtarget PlaceHalfPallet:=[[205,170,200],[0,0,1,0],[0,0,0,0],[9E+09,9E+09,9E+09,9E+09,9E+09,9E+09]];

    ! Liners
    CONST robtarget PickLiner:=[[400,270,100],[0,0,1,0],[0,0,0,0],[9E+09,9E+09,9E+09,9E+09,9E+09,9E+09]];
    CONST robtarget PlaceLiner:=[[400,300,210],[0,0,1,0],[0,0,0,0],[9E+09,9E+09,9E+09,9E+09,9E+09,9E+09]];

    !-----------------------------------------------------------------------
    ! Speeds and heights
    !-----------------------------------------------------------------------
    CONST speeddata TransitSpeed:=v1000;
    CONST speeddata ApproachSpeed:=v300;

    ! Height of every station (world)
    CONST num ConveyorsHeight:=768;
    CONST num TableHeight:=770;
    CONST num LinerStandHeight:=500;
    CONST num EuroPalletHeight:=144;
    CONST num HalfPalletHeight:=144;

    CONST num Box1Height:=200;
    CONST num Box2Height:=200;

    ! Heights for the approach points
    CONST num TransitHeight:=1100;
    CONST num PalletOffsetHeight:=250;
    CONST num MinApproachHeight:=250;

    ! Station identifiers for ApproachHeight
    CONST num StationConveyor1:=1;
    CONST num StationConveyor2:=2;
    CONST num StationTable:=3;
    CONST num StationLinerStand:=4;
    CONST num StationHalfPallet:=5;
    CONST num StationEuroPallet:=6;

    !-----------------------------------------------------------------------
    ! Vacuum gripper
    !-----------------------------------------------------------------------
    CONST num VacuumTime:=1;
    CONST bool CupsAllOn{6}:=[TRUE,TRUE,TRUE,TRUE,TRUE,TRUE];
    CONST bool CupsAllOff{6}:=[FALSE,FALSE,FALSE,FALSE,FALSE,FALSE];
    CONST bool CupsBox2On{6}:=[FALSE,FALSE,FALSE,TRUE,FALSE,FALSE];
    VAR signaldo cupSignals{6};

    !-----------------------------------------------------------------------
    ! Box selection
    !-----------------------------------------------------------------------
    CONST num Box1:=1;
    CONST num Box2:=2;
    ! Last box handled, to alternate box 1 and box 2
    VAR num lastBox:=Box2;

    !-----------------------------------------------------------------------
    ! Box 1 state machine parameters and variables
    !-----------------------------------------------------------------------
    CONST num Box1Pos1:=1;
    CONST num Box1Pos2:=2;
    CONST num Box1Pos3:=3;
    CONST num Box1Pos4:=4;
    CONST num Box1Pos5:=5;
    CONST num Box1LastPos:=6;
    CONST num Box1MaxLayers:=2;
    ! Distance between boxes in the row of 4 and in the row of 2
    CONST num EuroRow4Offset:=250;
    CONST num EuroRow2Offset:=500;

    VAR num box1State:=1;
    VAR num box1Layer:=1;
    VAR bool euroPalletFull:=FALSE;

    ! Euro pallet replaced by the operator: interrupt and flag set by the TRAP
    VAR intnum euroReplacedInt;
    VAR bool euroPalletReplaced:=FALSE;

    !-----------------------------------------------------------------------
    ! Box 2 state machine parameters and variables (table)
    !-----------------------------------------------------------------------
    CONST num Box2Pos1:=1;
    CONST num Box2Pos2:=2;
    CONST num Box2Pos3:=3;
    CONST num Box2Pos4:=4;
    CONST num Box2Pos5:=5;
    CONST num Box2LastPos:=6;
    ! Distance between boxes 2 on the table
    CONST num Box2Offset:=130;

    VAR num box2State:=1;
    VAR bool tableFull:=FALSE;

    !-----------------------------------------------------------------------
    ! TransferStack parameters and variables (half pallet)
    !-----------------------------------------------------------------------
    CONST num BlockPos1:=1;
    CONST num BlockPos2:=2;
    CONST num BlockPos3:=3;
    CONST num BlockPos4:=4;
    CONST num Box2MaxLayers:=3;
    ! Distance between 3x2 blocks on the half pallet
    CONST num BlockOffsetX:=3*Box2Offset;
    CONST num BlockOffsetY:=2*Box2Offset;

    VAR num blockState:=1;
    VAR num box2Layer:=1;
    VAR bool halfPalletFull:=FALSE;

    ! Half pallet replaced by the operator: interrupt and flag set by the TRAP
    VAR intnum halfReplacedInt;
    VAR bool halfPalletReplaced:=FALSE;

    !-----------------------------------------------------------------------
    ! Liners parameters and variables
    !-----------------------------------------------------------------------
    CONST num TotalLiners:=10;
    CONST num LinerHeight:=10;

    VAR num linersLeft:=TotalLiners;
    ! Liner stack empty: warning to the operator, the robot keeps working
    VAR bool linerStackEmpty:=FALSE;
    ! Layer complete but the liner stack is empty: box 2 waits for the refill
    VAR bool linerMissing:=FALSE;

    ! Liners refilled by the operator: interrupt and flag set by the TRAP
    VAR intnum linersRefilledInt;
    VAR bool linersRefilled:=FALSE;

    !-----------------------------------------------------------------------
    ! Main: choose the box and check the operator signals
    !-----------------------------------------------------------------------
    PROC Main()

        InitSignals;
        VacuumControl CupsAllOff;
        SetDO DO_EuroPalletFull,0;
        SetDO DO_HalfPalletFull,0;
        SetDO DO_LinerStackEmpty,0;
        ! Connect an interrupt to DI_EuroPalletReplaced: EuroPalletReplacedTrap runs on every rising edge
        IDelete euroReplacedInt;
        CONNECT euroReplacedInt WITH EuroPalletReplacedTrap;
        ISignalDI DI_EuroPalletReplaced,1,euroReplacedInt;
        ! Connect an interrupt to DI_HalfPalletReplaced: HalfPalletReplacedTrap runs on every rising edge
        IDelete halfReplacedInt;
        CONNECT halfReplacedInt WITH HalfPalletReplacedTrap;
        ISignalDI DI_HalfPalletReplaced,1,halfReplacedInt;
        ! Connect an interrupt to DI_LinersRefilled: LinersRefilledTrap runs on every rising edge
        IDelete linersRefilledInt;
        CONNECT linersRefilledInt WITH LinersRefilledTrap;
        ISignalDI DI_LinersRefilled,1,linersRefilledInt;
        GripLoad load0;
        MoveAbsJ Home,v100,fine,toolVacuum;

        WHILE TRUE DO

            ! Alternate box 1 and box 2 when both are ready
            IF Box1Ready() AND ((NOT Box2Ready()) OR lastBox=Box2) THEN
                ProcessBox1;
            ELSEIF Box2Ready() THEN
                ProcessBox2;
            ENDIF

            ! Euro pallet replaced (flag set by the TRAP): back to layer 1
            IF euroPalletReplaced THEN
                euroPalletReplaced:=FALSE;
                box1Layer:=1;
                ! Not necessary but safe
                box1State:=Box1Pos1;
                euroPalletFull:=FALSE;
            ENDIF

            ! Half pallet replaced (flag set by the TRAP): layer 1 first, then the waiting block
            IF halfPalletReplaced THEN
                halfPalletReplaced:=FALSE;
                box2Layer:=1;
                blockState:=BlockPos1;
                halfPalletFull:=FALSE;
                IF tableFull THEN
                    TransferStack;
                    tableFull:=FALSE;
                ENDIF
            ENDIF

            ! Liners refilled (flag set by the TRAP): reload the counter, then the missing liner and the waiting block
            IF linersRefilled THEN
                linersRefilled:=FALSE;
                linersLeft:=TotalLiners;
                linerStackEmpty:=FALSE;
                IF linerMissing THEN
                    linerMissing:=FALSE;
                    PlaceLayerLiner;
                    IF tableFull THEN
                        TransferStack;
                        tableFull:=FALSE;
                    ENDIF
                ENDIF
            ENDIF
            WaitTime 0.1;
        ENDWHILE
    ENDPROC

    !-----------------------------------------------------------------------
    ! Interrupts: operator buttons (pallet replaced, liners refilled)
    !-----------------------------------------------------------------------
    TRAP EuroPalletReplacedTrap
        ! Only considered if the pallet is already full to prevent false positives
        IF euroPalletFull THEN
            ! Light off at once, even while the robot moves: the operator instantly sees the press was accepted
            SetDO DO_EuroPalletFull,0;
            ! Main sets layer 1 when the robot is free (no motion in a TRAP)
            euroPalletReplaced:=TRUE;
        ENDIF
    ENDTRAP

    TRAP HalfPalletReplacedTrap
        ! Only considered if the pallet is already full to prevent false positives
        IF halfPalletFull THEN
            ! Light off at once, even while the robot moves: the operator instantly sees the press was accepted
            SetDO DO_HalfPalletFull,0;
            ! Main sets layer 1 and moves the waiting block (no motion in a TRAP)
            halfPalletReplaced:=TRUE;
        ENDIF
    ENDTRAP

    TRAP LinersRefilledTrap
        ! Only if the stack is empty, to prevent false positives
        IF linerStackEmpty THEN
            ! Light off at once, even while the robot moves: the operator instantly sees the press was accepted
            SetDO DO_LinerStackEmpty,0;
            ! Main reloads the counter, then places the missing liner and block (no motion in a TRAP)
            linersRefilled:=TRUE;
        ENDIF
    ENDTRAP

    !-----------------------------------------------------------------------
    ! Box ready to be handled
    !-----------------------------------------------------------------------
    FUNC bool Box1Ready()
        ! Box 1 waiting on conveyor 1 and room on the Euro pallet
        RETURN (DI_Box1Arrived=1) AND (NOT euroPalletFull);
    ENDFUNC

    FUNC bool Box2Ready()
        ! Box 2 waiting on conveyor 2 and room on the table
        RETURN (DI_Box2Arrived=1) AND (NOT tableFull);
    ENDFUNC

    !-----------------------------------------------------------------------
    ! Box 1 state machine: conveyor 1 to the Euro pallet
    !-----------------------------------------------------------------------
    PROC ProcessBox1()
        ! Z of the current layer on the Euro pallet
        VAR num layerZ;

        ApproachPoint PickConveyor1,wobjConveyor1,CupsAllOn,loadBox1,ApproachHeight(StationConveyor1);

        layerZ:=(box1Layer-1)*Box1Height;
        TEST box1State
        CASE Box1Pos1:
            ApproachPoint Offs(PlaceEuroRow4,0,0,layerZ),wobjEuroPallet,CupsAllOff,load0,ApproachHeight(StationEuroPallet);
            box1State:=Box1Pos2;
        CASE Box1Pos2:
            ApproachPoint Offs(PlaceEuroRow4,EuroRow4Offset,0,layerZ),wobjEuroPallet,CupsAllOff,load0,ApproachHeight(StationEuroPallet);
            box1State:=Box1Pos3;
        CASE Box1Pos3:
            ApproachPoint Offs(PlaceEuroRow4,2*EuroRow4Offset,0,layerZ),wobjEuroPallet,CupsAllOff,load0,ApproachHeight(StationEuroPallet);
            box1State:=Box1Pos4;
        CASE Box1Pos4:
            ApproachPoint Offs(PlaceEuroRow4,3*EuroRow4Offset,0,layerZ),wobjEuroPallet,CupsAllOff,load0,ApproachHeight(StationEuroPallet);
            box1State:=Box1Pos5;
        CASE Box1Pos5:
            ApproachPoint Offs(PlaceEuroRow2,0,0,layerZ),wobjEuroPallet,CupsAllOff,load0,ApproachHeight(StationEuroPallet);
            box1State:=Box1LastPos;
        CASE Box1LastPos:
            ApproachPoint Offs(PlaceEuroRow2,EuroRow2Offset,0,layerZ),wobjEuroPallet,CupsAllOff,load0,ApproachHeight(StationEuroPallet);
            IF box1Layer=Box1MaxLayers THEN
                euroPalletFull:=TRUE;
                SetDO DO_EuroPalletFull,1;
                TPWrite "Euro pallet full: replace it, then press the Euro pallet replaced button";
            ELSE
                Incr box1Layer;
            ENDIF
            box1State:=Box1Pos1;
        DEFAULT:
            box1State:=Box1Pos1;
        ENDTEST
        lastBox:=Box1;
    ENDPROC

    !-----------------------------------------------------------------------
    ! Box 2 state machine: conveyor 2 to the table
    !-----------------------------------------------------------------------
    PROC ProcessBox2()

        ApproachPoint PickConveyor2,wobjConveyor2,CupsBox2On,loadBox2,ApproachHeight(StationConveyor2);

        ! Far row (y=130) first and x from high to low: the box carried never crosses the boxes already placed
        TEST box2State
        CASE Box2Pos1:
            ApproachPoint Offs(PlaceTable,2*Box2Offset,Box2Offset,0),wobjTable,CupsAllOff,load0,ApproachHeight(StationTable);
            box2State:=Box2Pos2;
        CASE Box2Pos2:
            ApproachPoint Offs(PlaceTable,Box2Offset,Box2Offset,0),wobjTable,CupsAllOff,load0,ApproachHeight(StationTable);
            box2State:=Box2Pos3;
        CASE Box2Pos3:
            ApproachPoint Offs(PlaceTable,0,Box2Offset,0),wobjTable,CupsAllOff,load0,ApproachHeight(StationTable);
            box2State:=Box2Pos4;
        CASE Box2Pos4:
            ApproachPoint Offs(PlaceTable,2*Box2Offset,0,0),wobjTable,CupsAllOff,load0,ApproachHeight(StationTable);
            box2State:=Box2Pos5;
        CASE Box2Pos5:
            ApproachPoint Offs(PlaceTable,Box2Offset,0,0),wobjTable,CupsAllOff,load0,ApproachHeight(StationTable);
            box2State:=Box2LastPos;
        CASE Box2LastPos:
            ApproachPoint Offs(PlaceTable,0,0,0),wobjTable,CupsAllOff,load0,ApproachHeight(StationTable);
            IF halfPalletFull OR linerMissing THEN
                tableFull:=TRUE;
            ELSE
                TransferStack;
            ENDIF
            box2State:=Box2Pos1;
        DEFAULT:
            box2State:=Box2Pos1;
        ENDTEST
        lastBox:=Box2;
    ENDPROC

    !-----------------------------------------------------------------------
    ! Box 2: move the 3x2 block from the table to the half pallet
    !-----------------------------------------------------------------------
    PROC TransferStack()
        ! Z of the current layer on the half pallet (block and liner)
        VAR num layerZ;

        ! Pick all 6 boxes 2
        ApproachPoint PickTableStack,wobjTable,CupsAllOn,loadBox2Stack,ApproachHeight(StationTable);

        ! Place group of boxes
        layerZ:=HalfPalletLayerZ();
        TEST blockState
        CASE BlockPos1:
            ApproachPoint Offs(PlaceHalfPallet,0,BlockOffsetY,layerZ),wobjHalfPallet,CupsAllOff,load0,ApproachHeight(StationHalfPallet);
            blockState:=BlockPos2;
        CASE BlockPos2:
            ApproachPoint Offs(PlaceHalfPallet,BlockOffsetX,BlockOffsetY,layerZ),wobjHalfPallet,CupsAllOff,load0,ApproachHeight(StationHalfPallet);
            blockState:=BlockPos3;
        CASE BlockPos3:
            ApproachPoint Offs(PlaceHalfPallet,0,0,layerZ),wobjHalfPallet,CupsAllOff,load0,ApproachHeight(StationHalfPallet);
            blockState:=BlockPos4;
        CASE BlockPos4:
            ApproachPoint Offs(PlaceHalfPallet,BlockOffsetX,0,layerZ),wobjHalfPallet,CupsAllOff,load0,ApproachHeight(StationHalfPallet);
            IF box2Layer=Box2MaxLayers THEN
                halfPalletFull:=TRUE;
                SetDO DO_HalfPalletFull,1;
                TPWrite "Half pallet full: replace it, then press the half pallet replaced button";
            ELSEIF linerStackEmpty THEN
                linerMissing:=TRUE;
            ELSE
                PlaceLayerLiner;
            ENDIF
            blockState:=BlockPos1;
        DEFAULT:
            blockState:=BlockPos1;
        ENDTEST
    ENDPROC

    !-----------------------------------------------------------------------
    ! Liner on the layer just finished, then the next layer starts
    !-----------------------------------------------------------------------
    PROC PlaceLayerLiner()
        ApproachPoint Offs(PickLiner,0,0,-(TotalLiners-linersLeft)*LinerHeight),wobjLinerStack,CupsAllOn,loadLiner,ApproachHeight(StationLinerStand);
        ApproachPoint Offs(PlaceLiner,0,0,HalfPalletLayerZ()),wobjHalfPallet,CupsAllOff,load0,ApproachHeight(StationHalfPallet);
        Incr box2Layer;
        Decr linersLeft;
        IF linersLeft=0 THEN
            linerStackEmpty:=TRUE;
            SetDO DO_LinerStackEmpty,1;
            TPWrite "Liner stack empty: refill it, then press the liners refilled button";
        ENDIF
    ENDPROC

    !-----------------------------------------------------------------------
    ! Z of the current layer on the half pallet (block and liner)
    !-----------------------------------------------------------------------
    FUNC num HalfPalletLayerZ()
        ! One liner under every layer except the first one
        RETURN (box2Layer-1)*(Box2Height+LinerHeight);
    ENDFUNC

    !-----------------------------------------------------------------------
    ! Pick or place at a target: approach, vacuum, GripLoad and go up
    !-----------------------------------------------------------------------
    PROC ApproachPoint(robtarget target,PERS wobjdata wobj,bool cups{*},PERS loaddata load,num approachHeight)
        ! cups: cups on/off at the target, load: load after the target
        MoveJ Offs(target,0,0,approachHeight),TransitSpeed,z10,toolVacuum\WObj:=wobj;
        MoveL target,ApproachSpeed,fine,toolVacuum\WObj:=wobj;
        VacuumControl cups;
        GripLoad load;
        MoveL Offs(target,0,0,approachHeight),ApproachSpeed,z10,toolVacuum\WObj:=wobj;
    ENDPROC

    !-----------------------------------------------------------------------
    ! Calculation of approach heights (how much the robot goes up over the target)
    !-----------------------------------------------------------------------
    FUNC num ApproachHeight(num station)
        VAR num approachingHeight:=9E+09;
        TEST station
        CASE StationConveyor1:
            approachingHeight:=TransitHeight-ConveyorsHeight-Box1Height;
        CASE StationConveyor2:
            approachingHeight:=TransitHeight-ConveyorsHeight-Box2Height;
        CASE StationTable:
            approachingHeight:=TransitHeight-TableHeight-Box2Height;
        CASE StationLinerStand:
            approachingHeight:=TransitHeight-LinerStandHeight-linersLeft*LinerHeight;
        CASE StationHalfPallet:
            approachingHeight:=TransitHeight-HalfPalletHeight-HalfPalletLayerZ()-Box2Height-PalletOffsetHeight;
            IF approachingHeight<MinApproachHeight THEN
                approachingHeight:=MinApproachHeight;
            ENDIF
        CASE StationEuroPallet:
            approachingHeight:=TransitHeight-EuroPalletHeight-Box1Height*box1Layer-PalletOffsetHeight;
            IF approachingHeight<MinApproachHeight THEN
                approachingHeight:=MinApproachHeight;
            ENDIF
        DEFAULT:
            ! If another station is entered the robot will announce an error trying to reach 9E+09: Safety stop
        ENDTEST
        RETURN approachingHeight;
    ENDFUNC

    !-----------------------------------------------------------------------
    ! Assignment of logical cup signals with physical signals
    !-----------------------------------------------------------------------
    PROC InitSignals()
        ! Call it first: VacuumControl needs it
        AliasIO DO_Cup11,cupSignals{1};
        AliasIO DO_Cup12,cupSignals{2};
        AliasIO DO_Cup13,cupSignals{3};
        AliasIO DO_Cup21,cupSignals{4};
        AliasIO DO_Cup22,cupSignals{5};
        AliasIO DO_Cup23,cupSignals{6};
    ENDPROC

    !-----------------------------------------------------------------------
    ! Control of the vacuum of every cup
    !-----------------------------------------------------------------------
    PROC VacuumControl(bool cups{*})

        FOR i FROM 1 TO Dim(cups,1) DO
            IF cups{i} THEN
                SetDO cupSignals{i},1;
            ELSE
                SetDO cupSignals{i},0;
            ENDIF
        ENDFOR

        ! Robot stopped in position, wait for the vacuum
        WaitTime\InPos,VacuumTime;
    ENDPROC

ENDMODULE

--- Controller Data/Controler/SYSPAR/EIO.cfg ---
EIO:CFG_1.0:6:1::
#
EIO_SIGNAL:

      -Name "DO_Cup11" -SignalType "DO" -Label "Vacuum valve gripper"\
      -Category "Gripper"

      -Name "DI_Box1Arrived" -SignalType "DI" -Label "Box 1 sensor conveyor 1"\
      -Category "Conveyor"

      -Name "DI_Box2Arrived" -SignalType "DI" -Label "Box 2 sensor conveyor 2"\
      -Category "Conveyor"

      -Name "DI_EuroPalletReplaced" -SignalType "DI"\
      -Label "Operator confirms new euro pallet" -Category "Operator"

      -Name "DI_HalfPalletReplaced" -SignalType "DI"\
      -Label "Operator confirms new half pallet" -Category "Operator"

      -Name "AI_VacuumPressure" -SignalType "AI"\
      -Label "Vacuum pressure sensor (bar)" -Category "Gripper" -MaxLog 10

      -Name "DO_Cup12" -SignalType "DO" -Label "Vacuum valve gripper"\
      -Category "Gripper"

      -Name "DO_Cup13" -SignalType "DO" -Label "Vacuum valve gripper"\
      -Category "Gripper"

      -Name "DO_Cup21" -SignalType "DO" -Label "Vacuum valve gripper"\
      -Category "Gripper"

      -Name "DO_Cup22" -SignalType "DO" -Label "Vacuum valve gripper"\
      -Category "Gripper"

      -Name "DO_Cup23" -SignalType "DO" -Label "Vacuum valve gripper"\
      -Category "Gripper"

      -Name "DI_LinersRefilled" -SignalType "DI"\
      -Label "Indicates refilled liners" -Category "Liners"

      -Name "DO_EuroPalletFull" -SignalType "DO"

      -Name "DO_HalfPalletFull" -SignalType "DO"

      -Name "DO_LinerStackEmpty" -SignalType "DO"
